// 书籍分拣功能块主逻辑 - 使用上升沿检测提高鲁棒性
        // 1. 上升沿检测: 检测RFID传感器的上升沿（书籍到达时刻）
        Bin1_Trigger := RFID1 AND NOT LastRFID1;
        Bin2_Trigger := RFID2 AND NOT LastRFID2;
        Bin3_Trigger := RFID3 AND NOT LastRFID3;

        // 2. 电机控制逻辑: 任何RFID检测到书籍时启动电机
        Motor := RFID1 OR RFID2 OR RFID3;

        // 3. 分拣箱控制逻辑: 根据上升沿触发打开对应箱子，同一时间只有一个箱子打开
        // 优先级别: RFID1 > RFID2 > RFID3
        Bin1 := Bin1_Trigger AND NOT (Bin2_Trigger OR Bin3_Trigger);
        Bin2 := Bin2_Trigger AND NOT (Bin1_Trigger OR Bin3_Trigger);
        Bin3 := Bin3_Trigger AND NOT (Bin1_Trigger OR Bin2_Trigger);

        // 4. 更新上一周期状态
        LastRFID1 := RFID1;
        LastRFID2 := RFID2;
        LastRFID3 := RFID3;

        // 形式化属性验证断言
        // 属性1: 电机状态与RFID检测结果的一致性
        ASSERT((RFID1 OR RFID2 OR RFID3) = Motor);

        // 属性2: 同一时间最多只有一个箱子打开或全部关闭
        ASSERT(
          (Bin1 AND NOT Bin2 AND NOT Bin3) OR
          (Bin2 AND NOT Bin1 AND NOT Bin3) OR
          (Bin3 AND NOT Bin1 AND NOT Bin2) OR
          (NOT Bin1 AND NOT Bin2 AND NOT Bin3)
        );

        // 属性3: 无书籍时所有设备处于关闭状态
        ASSERT(
          (RFID1 OR RFID2 OR RFID3) OR
          (NOT Motor AND NOT Bin1 AND NOT Bin2 AND NOT Bin3)
        );
